(* PLC project g_bus_coupler_changeover_clean, Anonymous Benchmark Suite 1.0 *)
(* stored: creationDateTime 2026-09-02T00:00:00 *)

PROGRAM g_bus_coupler_changeover_clean
  VAR_INPUT
    incomer_a_healthy : BOOL;
    incomer_b_healthy : BOOL;
    maint : BOOL;
  END_VAR
  VAR_OUTPUT
    incomer_a : BOOL;
    incomer_b : BOOL;
    coupler : BOOL;
  END_VAR

(* LD diagram, written out as Structured Text *)
incomer_a := incomer_a_healthy;
incomer_b := incomer_b_healthy;
coupler := NOT incomer_a_healthy AND incomer_b_healthy;
END_PROGRAM

CONFIGURATION Config0
  RESOURCE Res0 ON PLC
    TASK tcyclic(INTERVAL := T#10ms, PRIORITY := 0);
    PROGRAM inst0 WITH tcyclic : g_bus_coupler_changeover_clean;
  END_RESOURCE
END_CONFIGURATION
